(* IEC 61131-3 sources: ArdisCVDCore/codesys/retired_hand_rolled_driver, 11 files *)

(* ---- ST_MfcChannelConfig.st ---- *)
TYPE ST_MfcChannelConfig :
STRUCT
    bSlaveAddr     : BYTE;
    sGasName       : STRING(8);
    rFullScaleSccm : REAL;
END_STRUCT
END_TYPE

(* ---- ST_MfcChannelState.st ---- *)
TYPE ST_MfcChannelState :
STRUCT
    iSubState       : INT;
    iRetryCount     : INT;
    wFaultCode      : WORD;
    xRegulating     : BOOL;
    xFaultActive    : BOOL;
    xCloseConfirmed : BOOL;
    rMeasuredSccm   : REAL;
END_STRUCT
END_TYPE

(* ---- F_MbReadFrame.st ---- *)
FUNCTION F_MbReadFrame : INT
VAR_INPUT
    bAddr : BYTE;
    wReg  : WORD;
END_VAR
VAR_IN_OUT
    aFrame : ARRAY[0..7] OF BYTE;
END_VAR
VAR
    wCrc : WORD;
END_VAR

aFrame[0] := bAddr;
aFrame[1] := BYTE#16#03;
aFrame[2] := WORD_TO_BYTE(SHR(wReg, 8));
aFrame[3] := WORD_TO_BYTE(wReg AND WORD#16#00FF);
aFrame[4] := BYTE#0;
aFrame[5] := BYTE#1;
wCrc := F_ModbusCrc16(iLen := 6, aData := aFrame);
aFrame[6] := WORD_TO_BYTE(wCrc AND WORD#16#00FF);
aFrame[7] := WORD_TO_BYTE(SHR(wCrc, 8));

F_MbReadFrame := 8;

(* ---- F_MbReadStep.st ---- *)
FUNCTION F_MbReadStep : INT
VAR_INPUT
    xReadDone   : BOOL;
    xReadError  : BOOL;
    udiReadSize : UDINT;
END_VAR
VAR_IN_OUT
    xReadExecute    : BOOL;
    xRetriggerArmed : BOOL;
    iRxAccum        : INT;
    iRxIdleScans    : INT;
END_VAR
VAR CONSTANT
    C_MAX_FRAME       : INT := 8;
    C_IDLE_SCAN_LIMIT : INT := 2;
    C_NODATA_LIMIT    : INT := 3;
END_VAR

IF xRetriggerArmed THEN
    xRetriggerArmed := FALSE;
    xReadExecute := TRUE;
    F_MbReadStep := 0;
    RETURN;
END_IF;

IF xReadError THEN
    xReadExecute := FALSE;
    F_MbReadStep := 2;
    RETURN;
END_IF;

IF NOT xReadDone THEN
    F_MbReadStep := 0;
    RETURN;
END_IF;

IF udiReadSize > UDINT#0 THEN
    iRxAccum := iRxAccum + UDINT_TO_INT(udiReadSize);
    iRxIdleScans := 0;
ELSE
    iRxIdleScans := iRxIdleScans + 1;
END_IF;

IF iRxAccum >= C_MAX_FRAME THEN
    xReadExecute := FALSE;
    F_MbReadStep := 1;
    RETURN;
END_IF;

IF (iRxAccum > 0) AND (iRxIdleScans >= C_IDLE_SCAN_LIMIT) THEN
    xReadExecute := FALSE;
    F_MbReadStep := 1;
    RETURN;
END_IF;

IF (iRxAccum = 0) AND (iRxIdleScans >= C_NODATA_LIMIT) THEN
    xReadExecute := FALSE;
    F_MbReadStep := 2;
    RETURN;
END_IF;

xReadExecute := FALSE;
xRetriggerArmed := TRUE;
F_MbReadStep := 0;

(* ---- F_MbRetryOrFault.st ---- *)
FUNCTION F_MbRetryOrFault : INT
VAR_INPUT
    iIssueState : INT;
    iFaultState : INT;
    iMaxRetries : INT;
END_VAR
VAR_IN_OUT
    iRetryCount : INT;
END_VAR

IF iRetryCount < iMaxRetries THEN
    iRetryCount := iRetryCount + 1;
    F_MbRetryOrFault := iIssueState;
ELSE
    iRetryCount := 0;
    F_MbRetryOrFault := iFaultState;
END_IF;

(* ---- F_MbValidateResponse.st ---- *)
FUNCTION F_MbValidateResponse : WORD
VAR_INPUT
    iSize        : INT;
    bExpectAddr  : BYTE;
    bExpectFunc  : BYTE;
    wExpectReg   : WORD;
    wExpectValue : WORD;
    xIsWrite     : BOOL;
END_VAR
VAR_IN_OUT
    aFrame : ARRAY[0..7] OF BYTE;
END_VAR
VAR_OUTPUT
    wReadValue : WORD;
END_VAR
VAR
    wCrcCalc   : WORD;
    wCrcRecv   : WORD;
    iExpectLen : INT;
END_VAR

wReadValue := WORD#0;

IF xIsWrite THEN
    iExpectLen := 8;
ELSE
    iExpectLen := 7;
END_IF;

IF (iSize <> iExpectLen) AND (iSize <> 5) THEN
    F_MbValidateResponse := WORD#5;
    RETURN;
END_IF;

wCrcCalc := F_ModbusCrc16(iLen := iSize - 2, aData := aFrame);
wCrcRecv := BYTE_TO_WORD(aFrame[iSize - 2]) OR SHL(BYTE_TO_WORD(aFrame[iSize - 1]), 8);
IF wCrcCalc <> wCrcRecv THEN
    F_MbValidateResponse := WORD#3;
    RETURN;
END_IF;

IF aFrame[0] <> bExpectAddr THEN
    F_MbValidateResponse := WORD#6;
    RETURN;
END_IF;

IF aFrame[1] = (bExpectFunc OR BYTE#16#80) THEN
    F_MbValidateResponse := WORD#4;
    RETURN;
END_IF;

IF aFrame[1] <> bExpectFunc THEN
    F_MbValidateResponse := WORD#7;
    RETURN;
END_IF;

IF xIsWrite THEN
    IF (aFrame[2] <> WORD_TO_BYTE(SHR(wExpectReg, 8))) OR
       (aFrame[3] <> WORD_TO_BYTE(wExpectReg AND WORD#16#00FF)) OR
       (aFrame[4] <> WORD_TO_BYTE(SHR(wExpectValue, 8))) OR
       (aFrame[5] <> WORD_TO_BYTE(wExpectValue AND WORD#16#00FF)) THEN
        F_MbValidateResponse := WORD#8;
        RETURN;
    END_IF;
ELSE
    wReadValue := SHL(BYTE_TO_WORD(aFrame[3]), 8) OR BYTE_TO_WORD(aFrame[4]);
END_IF;

F_MbValidateResponse := WORD#0;

(* ---- F_MbWriteFrame.st ---- *)
FUNCTION F_MbWriteFrame : INT
VAR_INPUT
    bAddr  : BYTE;
    wReg   : WORD;
    wValue : WORD;
END_VAR
VAR_IN_OUT
    aFrame : ARRAY[0..7] OF BYTE;
END_VAR
VAR
    wCrc : WORD;
END_VAR

aFrame[0] := bAddr;
aFrame[1] := BYTE#16#06;
aFrame[2] := WORD_TO_BYTE(SHR(wReg, 8));
aFrame[3] := WORD_TO_BYTE(wReg AND WORD#16#00FF);
aFrame[4] := WORD_TO_BYTE(SHR(wValue, 8));
aFrame[5] := WORD_TO_BYTE(wValue AND WORD#16#00FF);
wCrc := F_ModbusCrc16(iLen := 6, aData := aFrame);
aFrame[6] := WORD_TO_BYTE(wCrc AND WORD#16#00FF);
aFrame[7] := WORD_TO_BYTE(SHR(wCrc, 8));

F_MbWriteFrame := 8;

(* ---- F_ModbusCrc16.st ---- *)
FUNCTION F_ModbusCrc16 : WORD
VAR_INPUT
    iLen : INT;
END_VAR
VAR_IN_OUT
    aData : ARRAY[0..7] OF BYTE;
END_VAR
VAR
    wCrc : WORD;
    i    : INT;
    j    : INT;
END_VAR

wCrc := WORD#16#FFFF;
FOR i := 0 TO iLen - 1 DO
    wCrc := wCrc XOR BYTE_TO_WORD(aData[i]);
    FOR j := 0 TO 7 DO
        IF (wCrc AND WORD#16#0001) = WORD#16#0001 THEN
            wCrc := SHR(wCrc, 1) XOR WORD#16#A001;
        ELSE
            wCrc := SHR(wCrc, 1);
        END_IF;
    END_FOR;
END_FOR;

F_ModbusCrc16 := wCrc;

(* ---- FB_IncrementalPidOLD.st ---- *)
FUNCTION_BLOCK FB_IncrementalPid
VAR_INPUT
    xEnable       : BOOL;
    xReset        : BOOL;
    xDirectMode   : BOOL;
    rSetpoint     : REAL;
    rMeasured     : REAL;
    rKp           : REAL;
    rKi           : REAL;
    rKd           : REAL;
    rLowerLimit   : REAL;
    rUpperLimit   : REAL;
    rDirectValue  : REAL;
    rFlowCorrection     : REAL := 1.0;
    rPressureCorrection : REAL := 1.0;
    rTotalGasFlow       : REAL := 0.0;
    rCycleSeconds : REAL := 0.2;
END_VAR
VAR_OUTPUT
    rError  : REAL;
    rP      : REAL;
    rI      : REAL;
    rD      : REAL;
    rOutput : REAL;
END_VAR
VAR
    rIntegral      : REAL;
    rPreviousError : REAL;
    xInitialized   : BOOL;
    rMin           : REAL;
    rMax           : REAL;
    rFlowScale     : REAL;
    rPressureScale : REAL;
END_VAR

IF rLowerLimit <= rUpperLimit THEN
    rMin := rLowerLimit;
    rMax := rUpperLimit;
ELSE
    rMin := rUpperLimit;
    rMax := rLowerLimit;
END_IF;

rError := rMeasured - rSetpoint;

IF NOT xEnable THEN
    rP := 0.0;
    rI := 0.0;
    rD := 0.0;
    rOutput := rMin;
    rIntegral := 0.0;
    rPreviousError := rError;
    xInitialized := FALSE;
    RETURN;
END_IF;

IF xReset OR NOT xInitialized THEN
    rIntegral := 0.0;
    rPreviousError := rError;
    rOutput := rMin;
    xInitialized := TRUE;
END_IF;

rP := rKp * rError;

IF rCycleSeconds > 0.001 THEN
    rIntegral := rIntegral + rError * rCycleSeconds;
    rD := rKd * (rError - rPreviousError) / rCycleSeconds;
ELSE
    rD := 0.0;
END_IF;

IF (rFlowCorrection > 0.001) AND (rTotalGasFlow > 50.0) THEN
    IF rTotalGasFlow <= 1100.0 THEN
        rFlowScale := ((rTotalGasFlow - 50.0) / (1100.0 - 50.0)) * (rFlowCorrection - 1.0) + 1.0;
    ELSE
        rFlowScale := rFlowCorrection;
    END_IF;

    IF rFlowScale > 0.001 THEN
        rP := rP / rFlowScale;
        rD := rD / rFlowScale;
    END_IF;
END_IF;

IF (rPressureCorrection > 0.001) AND (rMeasured > 10.0) THEN
    IF rMeasured < 500.0 THEN
        rPressureScale := ((rMeasured - 10.0) / (500.0 - 10.0)) * (rPressureCorrection - 1.0) + 1.0;
    ELSE
        rPressureScale := rPressureCorrection;
    END_IF;

    IF rPressureScale > 0.001 THEN
        rP := rP / rPressureScale;
        rD := rD / rPressureScale;
    END_IF;
END_IF;

IF rIntegral > 1000000.0 THEN
    rIntegral := 1000000.0;
ELSIF rIntegral < -1000000.0 THEN
    rIntegral := -1000000.0;
END_IF;

rI := rKi * rIntegral;
rPreviousError := rError;

IF xDirectMode THEN
    rOutput := rDirectValue;
ELSE
    rOutput := rOutput + rP + rI + rD;
END_IF;

IF rOutput > rMax THEN
    rOutput := rMax;
ELSIF rOutput < rMin THEN
    rOutput := rMin;
END_IF;

(* ---- FB_MfcModbusMaster.st ---- *)
FUNCTION_BLOCK FB_MfcModbusMaster
VAR_INPUT
    xEnable        : BOOL;
    udiPort        : UDINT := 4;
    udiBaudrate    : UDINT := 19200;
    arSetpointSccm : ARRAY[0..5] OF REAL;
END_VAR
VAR_OUTPUT
    xBusOpen         : BOOL;
    udiSweepCounter  : UDINT;
    arMeasuredSccm   : ARRAY[0..5] OF REAL;
    axRegulating     : ARRAY[0..5] OF BOOL;
    axFaultActive    : ARRAY[0..5] OF BOOL;
    axCloseConfirmed : ARRAY[0..5] OF BOOL;
    awFaultCode      : ARRAY[0..5] OF WORD;
END_VAR
VAR CONSTANT
    C_REG_MODE         : WORD := 2;
    C_REG_SETPOINT     : WORD := 4;
    C_REG_MEASURED     : WORD := 5;
    C_REG_RAMPTIME     : WORD := 19;
    C_REG_RAMPSTEP     : WORD := 20;
    C_REG_RAMPEN       : WORD := 21;
    C_MODE_REGULATE    : WORD := 19;
    C_MODE_CLOSE       : WORD := 10;
    C_RAMPTIME_DEFAULT : WORD := 200;
    C_RAMPSTEP_DEFAULT : WORD := 10;
    C_RAMPEN_DEFAULT   : WORD := 1;
    C_FUNC_READ        : BYTE := 16#03;
    C_FUNC_WRITE       : BYTE := 16#06;
    C_MAX_RETRIES      : INT := 2;
    C_OPEN_RETRY_TICKS : UDINT := 40;
    C_IO_TIMEOUT_US    : UDINT := 100000;
END_VAR
VAR
    aCfg        : ARRAY[0..5] OF ST_MfcChannelConfig;
    xConfigInit : BOOL;

    aCh : ARRAY[0..5] OF ST_MfcChannelState;

    iBusState         : INT;
    iChannel          : INT;
    hCom              : CAA.HANDLE;
    udiOpenRetryTicks : UDINT;

    fbOpen  : COM.Open;
    fbWrite : COM.Write;
    fbRead  : COM.Read;
    aParams : ARRAY[1..7] OF COM.PARAMETER;
    xOpenExecute  : BOOL;
    xWriteExecute : BOOL;
    xReadExecute  : BOOL;

    aTx     : ARRAY[0..7] OF BYTE;
    aRx     : ARRAY[0..7] OF BYTE;
    iRxSize : INT;

    iRxAccum         : INT;
    iRxIdleScans     : INT;
    xRxRetriggerArmed: BOOL;
    iRxOffset        : INT;
    iAccumStatus     : INT;

    bPendingAddr    : BYTE;
    wPendingReg     : WORD;
    wPendingValue   : WORD;

    wValidateResult : WORD;
    wReadValue      : WORD;
    rRaw            : REAL;
    iRawSetpoint    : INT;

    i : INT;
END_VAR

IF NOT xConfigInit THEN
    aCfg[0].bSlaveAddr := BYTE#1; aCfg[0].sGasName := 'H2';  aCfg[0].rFullScaleSccm := 1000.0;
    aCfg[1].bSlaveAddr := BYTE#2; aCfg[1].sGasName := 'CH4'; aCfg[1].rFullScaleSccm := 100.0;
    aCfg[2].bSlaveAddr := BYTE#3; aCfg[2].sGasName := 'O2';  aCfg[2].rFullScaleSccm := 50.0;
    aCfg[3].bSlaveAddr := BYTE#4; aCfg[3].sGasName := 'N2';  aCfg[3].rFullScaleSccm := 1000.0;
    aCfg[4].bSlaveAddr := BYTE#5; aCfg[4].sGasName := 'Ar';  aCfg[4].rFullScaleSccm := 10.0;
    aCfg[5].bSlaveAddr := BYTE#6; aCfg[5].sGasName := 'H22'; aCfg[5].rFullScaleSccm := 1000.0;
    xConfigInit := TRUE;
END_IF;

IF NOT xEnable THEN
    FOR i := 0 TO 5 DO
        IF (aCh[i].iSubState <> 900) AND (aCh[i].iSubState <> 901) AND (aCh[i].iSubState <> 902) THEN
            aCh[i].iSubState := 900;
            aCh[i].iRetryCount := 0;
        END_IF;
    END_FOR;
END_IF;

aParams[1].udiParameterId := COM.CAA_Parameter_Constants.udiPort;
aParams[1].udiValue := udiPort;
aParams[2].udiParameterId := COM.CAA_Parameter_Constants.udiBaudrate;
aParams[2].udiValue := udiBaudrate;
aParams[3].udiParameterId := COM.CAA_Parameter_Constants.udiParity;
aParams[3].udiValue := 2;
aParams[4].udiParameterId := COM.CAA_Parameter_Constants.udiStopBits;
aParams[4].udiValue := 0;
aParams[5].udiParameterId := COM.CAA_Parameter_Constants.udiTimeout;
aParams[5].udiValue := 200000;
aParams[6].udiParameterId := COM.CAA_Parameter_Constants.udiByteSize;
aParams[6].udiValue := 8;
aParams[7].udiParameterId := COM.CAA_Parameter_Constants.udiBinary;
aParams[7].udiValue := 1;

CASE iBusState OF

    0:
        xOpenExecute := TRUE;
        xBusOpen := FALSE;
        IF fbOpen.xDone THEN
            hCom := fbOpen.hCom;
            xOpenExecute := FALSE;
            xBusOpen := TRUE;
            iChannel := 0;
            FOR i := 0 TO 5 DO
                IF xEnable THEN
                    aCh[i].iSubState := 100;
                ELSE
                    aCh[i].iSubState := 900;
                END_IF;
                aCh[i].iRetryCount := 0;
            END_FOR;
            iBusState := 10;
        ELSIF fbOpen.xError THEN
            xOpenExecute := FALSE;
            udiOpenRetryTicks := 0;
            iBusState := 5;
        END_IF;

    5:
        xBusOpen := FALSE;
        udiOpenRetryTicks := udiOpenRetryTicks + 1;
        IF udiOpenRetryTicks >= C_OPEN_RETRY_TICKS THEN
            iBusState := 0;
        END_IF;

    10:
        CASE aCh[iChannel].iSubState OF

            100:
                bPendingAddr := aCfg[iChannel].bSlaveAddr;
                wPendingReg := C_REG_RAMPTIME;
                wPendingValue := C_RAMPTIME_DEFAULT;
                F_MbWriteFrame(bAddr := bPendingAddr, wReg := wPendingReg, wValue := wPendingValue, aFrame := aTx);
                xWriteExecute := TRUE;
                aCh[iChannel].iSubState := 101;

            101:
                IF fbWrite.xDone THEN
                    xWriteExecute := FALSE;
                    xReadExecute := TRUE;
                    iRxAccum := 0;
                    iRxIdleScans := 0;
                    xRxRetriggerArmed := FALSE;
                    aCh[iChannel].iSubState := 102;
                ELSIF fbWrite.xError THEN
                    xWriteExecute := FALSE;
                    aCh[iChannel].wFaultCode := WORD#1;
                    aCh[iChannel].iSubState := F_MbRetryOrFault(iIssueState := 100, iFaultState := 900, iMaxRetries := C_MAX_RETRIES, iRetryCount := aCh[iChannel].iRetryCount);
                END_IF;

            102:
                iAccumStatus := F_MbReadStep(xReadDone := fbRead.xDone, xReadError := fbRead.xError, udiReadSize := fbRead.szSize,
                    xReadExecute := xReadExecute, xRetriggerArmed := xRxRetriggerArmed, iRxAccum := iRxAccum, iRxIdleScans := iRxIdleScans);
                IF iAccumStatus = 1 THEN
                    iRxSize := iRxAccum;
                    wValidateResult := F_MbValidateResponse(iSize := iRxSize, bExpectAddr := bPendingAddr, bExpectFunc := C_FUNC_WRITE,
                        wExpectReg := wPendingReg, wExpectValue := wPendingValue, xIsWrite := TRUE, aFrame := aRx, wReadValue => wReadValue);
                    IF wValidateResult = WORD#0 THEN
                        aCh[iChannel].iRetryCount := 0;
                        aCh[iChannel].iSubState := 110;
                    ELSE
                        aCh[iChannel].wFaultCode := wValidateResult;
                        aCh[iChannel].iSubState := F_MbRetryOrFault(iIssueState := 100, iFaultState := 900, iMaxRetries := C_MAX_RETRIES, iRetryCount := aCh[iChannel].iRetryCount);
                    END_IF;
                ELSIF iAccumStatus = 2 THEN
                    aCh[iChannel].wFaultCode := WORD#2;
                    aCh[iChannel].iSubState := F_MbRetryOrFault(iIssueState := 100, iFaultState := 900, iMaxRetries := C_MAX_RETRIES, iRetryCount := aCh[iChannel].iRetryCount);
                END_IF;

            110:
                bPendingAddr := aCfg[iChannel].bSlaveAddr;
                wPendingReg := C_REG_RAMPSTEP;
                wPendingValue := C_RAMPSTEP_DEFAULT;
                F_MbWriteFrame(bAddr := bPendingAddr, wReg := wPendingReg, wValue := wPendingValue, aFrame := aTx);
                xWriteExecute := TRUE;
                aCh[iChannel].iSubState := 111;

            111:
                IF fbWrite.xDone THEN
                    xWriteExecute := FALSE;
                    xReadExecute := TRUE;
                    iRxAccum := 0;
                    iRxIdleScans := 0;
                    xRxRetriggerArmed := FALSE;
                    aCh[iChannel].iSubState := 112;
                ELSIF fbWrite.xError THEN
                    xWriteExecute := FALSE;
                    aCh[iChannel].wFaultCode := WORD#1;
                    aCh[iChannel].iSubState := F_MbRetryOrFault(iIssueState := 110, iFaultState := 900, iMaxRetries := C_MAX_RETRIES, iRetryCount := aCh[iChannel].iRetryCount);
                END_IF;

            112:
                iAccumStatus := F_MbReadStep(xReadDone := fbRead.xDone, xReadError := fbRead.xError, udiReadSize := fbRead.szSize,
                    xReadExecute := xReadExecute, xRetriggerArmed := xRxRetriggerArmed, iRxAccum := iRxAccum, iRxIdleScans := iRxIdleScans);
                IF iAccumStatus = 1 THEN
                    iRxSize := iRxAccum;
                    wValidateResult := F_MbValidateResponse(iSize := iRxSize, bExpectAddr := bPendingAddr, bExpectFunc := C_FUNC_WRITE,
                        wExpectReg := wPendingReg, wExpectValue := wPendingValue, xIsWrite := TRUE, aFrame := aRx, wReadValue => wReadValue);
                    IF wValidateResult = WORD#0 THEN
                        aCh[iChannel].iRetryCount := 0;
                        aCh[iChannel].iSubState := 120;
                    ELSE
                        aCh[iChannel].wFaultCode := wValidateResult;
                        aCh[iChannel].iSubState := F_MbRetryOrFault(iIssueState := 110, iFaultState := 900, iMaxRetries := C_MAX_RETRIES, iRetryCount := aCh[iChannel].iRetryCount);
                    END_IF;
                ELSIF iAccumStatus = 2 THEN
                    aCh[iChannel].wFaultCode := WORD#2;
                    aCh[iChannel].iSubState := F_MbRetryOrFault(iIssueState := 110, iFaultState := 900, iMaxRetries := C_MAX_RETRIES, iRetryCount := aCh[iChannel].iRetryCount);
                END_IF;

            120:
                bPendingAddr := aCfg[iChannel].bSlaveAddr;
                wPendingReg := C_REG_RAMPEN;
                wPendingValue := C_RAMPEN_DEFAULT;
                F_MbWriteFrame(bAddr := bPendingAddr, wReg := wPendingReg, wValue := wPendingValue, aFrame := aTx);
                xWriteExecute := TRUE;
                aCh[iChannel].iSubState := 121;

            121:
                IF fbWrite.xDone THEN
                    xWriteExecute := FALSE;
                    xReadExecute := TRUE;
                    iRxAccum := 0;
                    iRxIdleScans := 0;
                    xRxRetriggerArmed := FALSE;
                    aCh[iChannel].iSubState := 122;
                ELSIF fbWrite.xError THEN
                    xWriteExecute := FALSE;
                    aCh[iChannel].wFaultCode := WORD#1;
                    aCh[iChannel].iSubState := F_MbRetryOrFault(iIssueState := 120, iFaultState := 900, iMaxRetries := C_MAX_RETRIES, iRetryCount := aCh[iChannel].iRetryCount);
                END_IF;

            122:
                iAccumStatus := F_MbReadStep(xReadDone := fbRead.xDone, xReadError := fbRead.xError, udiReadSize := fbRead.szSize,
                    xReadExecute := xReadExecute, xRetriggerArmed := xRxRetriggerArmed, iRxAccum := iRxAccum, iRxIdleScans := iRxIdleScans);
                IF iAccumStatus = 1 THEN
                    iRxSize := iRxAccum;
                    wValidateResult := F_MbValidateResponse(iSize := iRxSize, bExpectAddr := bPendingAddr, bExpectFunc := C_FUNC_WRITE,
                        wExpectReg := wPendingReg, wExpectValue := wPendingValue, xIsWrite := TRUE, aFrame := aRx, wReadValue => wReadValue);
                    IF wValidateResult = WORD#0 THEN
                        aCh[iChannel].iRetryCount := 0;
                        aCh[iChannel].iSubState := 130;
                    ELSE
                        aCh[iChannel].wFaultCode := wValidateResult;
                        aCh[iChannel].iSubState := F_MbRetryOrFault(iIssueState := 120, iFaultState := 900, iMaxRetries := C_MAX_RETRIES, iRetryCount := aCh[iChannel].iRetryCount);
                    END_IF;
                ELSIF iAccumStatus = 2 THEN
                    aCh[iChannel].wFaultCode := WORD#2;
                    aCh[iChannel].iSubState := F_MbRetryOrFault(iIssueState := 120, iFaultState := 900, iMaxRetries := C_MAX_RETRIES, iRetryCount := aCh[iChannel].iRetryCount);
                END_IF;

            130:
                bPendingAddr := aCfg[iChannel].bSlaveAddr;
                wPendingReg := C_REG_MODE;
                wPendingValue := C_MODE_REGULATE;
                F_MbWriteFrame(bAddr := bPendingAddr, wReg := wPendingReg, wValue := wPendingValue, aFrame := aTx);
                xWriteExecute := TRUE;
                aCh[iChannel].iSubState := 131;

            131:
                IF fbWrite.xDone THEN
                    xWriteExecute := FALSE;
                    xReadExecute := TRUE;
                    iRxAccum := 0;
                    iRxIdleScans := 0;
                    xRxRetriggerArmed := FALSE;
                    aCh[iChannel].iSubState := 132;
                ELSIF fbWrite.xError THEN
                    xWriteExecute := FALSE;
                    aCh[iChannel].wFaultCode := WORD#1;
                    aCh[iChannel].iSubState := F_MbRetryOrFault(iIssueState := 130, iFaultState := 900, iMaxRetries := C_MAX_RETRIES, iRetryCount := aCh[iChannel].iRetryCount);
                END_IF;

            132:
                iAccumStatus := F_MbReadStep(xReadDone := fbRead.xDone, xReadError := fbRead.xError, udiReadSize := fbRead.szSize,
                    xReadExecute := xReadExecute, xRetriggerArmed := xRxRetriggerArmed, iRxAccum := iRxAccum, iRxIdleScans := iRxIdleScans);
                IF iAccumStatus = 1 THEN
                    iRxSize := iRxAccum;
                    wValidateResult := F_MbValidateResponse(iSize := iRxSize, bExpectAddr := bPendingAddr, bExpectFunc := C_FUNC_WRITE,
                        wExpectReg := wPendingReg, wExpectValue := wPendingValue, xIsWrite := TRUE, aFrame := aRx, wReadValue => wReadValue);
                    IF wValidateResult = WORD#0 THEN
                        aCh[iChannel].iRetryCount := 0;
                        aCh[iChannel].wFaultCode := WORD#0;
                        aCh[iChannel].xFaultActive := FALSE;
                        aCh[iChannel].xCloseConfirmed := FALSE;
                        aCh[iChannel].xRegulating := TRUE;
                        aCh[iChannel].iSubState := 200;
                    ELSE
                        aCh[iChannel].wFaultCode := wValidateResult;
                        aCh[iChannel].iSubState := F_MbRetryOrFault(iIssueState := 130, iFaultState := 900, iMaxRetries := C_MAX_RETRIES, iRetryCount := aCh[iChannel].iRetryCount);
                    END_IF;
                ELSIF iAccumStatus = 2 THEN
                    aCh[iChannel].wFaultCode := WORD#2;
                    aCh[iChannel].iSubState := F_MbRetryOrFault(iIssueState := 130, iFaultState := 900, iMaxRetries := C_MAX_RETRIES, iRetryCount := aCh[iChannel].iRetryCount);
                END_IF;

            200:
                rRaw := arSetpointSccm[iChannel] / aCfg[iChannel].rFullScaleSccm * 10000.0;
                IF rRaw < 0.0 THEN
                    rRaw := 0.0;
                END_IF;
                iRawSetpoint := REAL_TO_INT(rRaw + 0.5);
                IF iRawSetpoint > 10000 THEN
                    iRawSetpoint := 10000;
                ELSIF iRawSetpoint < 0 THEN
                    iRawSetpoint := 0;
                END_IF;

                bPendingAddr := aCfg[iChannel].bSlaveAddr;
                wPendingReg := C_REG_SETPOINT;
                wPendingValue := INT_TO_WORD(iRawSetpoint);
                F_MbWriteFrame(bAddr := bPendingAddr, wReg := wPendingReg, wValue := wPendingValue, aFrame := aTx);
                xWriteExecute := TRUE;
                aCh[iChannel].iSubState := 201;

            201:
                IF fbWrite.xDone THEN
                    xWriteExecute := FALSE;
                    xReadExecute := TRUE;
                    iRxAccum := 0;
                    iRxIdleScans := 0;
                    xRxRetriggerArmed := FALSE;
                    aCh[iChannel].iSubState := 202;
                ELSIF fbWrite.xError THEN
                    xWriteExecute := FALSE;
                    aCh[iChannel].wFaultCode := WORD#1;
                    aCh[iChannel].iSubState := F_MbRetryOrFault(iIssueState := 200, iFaultState := 900, iMaxRetries := C_MAX_RETRIES, iRetryCount := aCh[iChannel].iRetryCount);
                END_IF;

            202:
                iAccumStatus := F_MbReadStep(xReadDone := fbRead.xDone, xReadError := fbRead.xError, udiReadSize := fbRead.szSize,
                    xReadExecute := xReadExecute, xRetriggerArmed := xRxRetriggerArmed, iRxAccum := iRxAccum, iRxIdleScans := iRxIdleScans);
                IF iAccumStatus = 1 THEN
                    iRxSize := iRxAccum;
                    wValidateResult := F_MbValidateResponse(iSize := iRxSize, bExpectAddr := bPendingAddr, bExpectFunc := C_FUNC_WRITE,
                        wExpectReg := wPendingReg, wExpectValue := wPendingValue, xIsWrite := TRUE, aFrame := aRx, wReadValue => wReadValue);
                    IF wValidateResult = WORD#0 THEN
                        aCh[iChannel].iRetryCount := 0;
                        aCh[iChannel].iSubState := 210;
                    ELSE
                        aCh[iChannel].wFaultCode := wValidateResult;
                        aCh[iChannel].iSubState := F_MbRetryOrFault(iIssueState := 200, iFaultState := 900, iMaxRetries := C_MAX_RETRIES, iRetryCount := aCh[iChannel].iRetryCount);
                    END_IF;
                ELSIF iAccumStatus = 2 THEN
                    aCh[iChannel].wFaultCode := WORD#2;
                    aCh[iChannel].iSubState := F_MbRetryOrFault(iIssueState := 200, iFaultState := 900, iMaxRetries := C_MAX_RETRIES, iRetryCount := aCh[iChannel].iRetryCount);
                END_IF;

            210:
                bPendingAddr := aCfg[iChannel].bSlaveAddr;
                wPendingReg := C_REG_MEASURED;
                F_MbReadFrame(bAddr := bPendingAddr, wReg := wPendingReg, aFrame := aTx);
                xReadExecute := TRUE;
                iRxAccum := 0;
                iRxIdleScans := 0;
                xRxRetriggerArmed := FALSE;
                aCh[iChannel].iSubState := 211;

            211:
                iAccumStatus := F_MbReadStep(xReadDone := fbRead.xDone, xReadError := fbRead.xError, udiReadSize := fbRead.szSize,
                    xReadExecute := xReadExecute, xRetriggerArmed := xRxRetriggerArmed, iRxAccum := iRxAccum, iRxIdleScans := iRxIdleScans);
                IF iAccumStatus = 1 THEN
                    iRxSize := iRxAccum;
                    wValidateResult := F_MbValidateResponse(iSize := iRxSize, bExpectAddr := bPendingAddr, bExpectFunc := C_FUNC_READ,
                        wExpectReg := wPendingReg, wExpectValue := WORD#0, xIsWrite := FALSE, aFrame := aRx, wReadValue => wReadValue);
                    IF wValidateResult = WORD#0 THEN
                        aCh[iChannel].iRetryCount := 0;
                        aCh[iChannel].rMeasuredSccm := UINT_TO_REAL(WORD_TO_UINT(wReadValue)) / 10000.0 * aCfg[iChannel].rFullScaleSccm;
                        aCh[iChannel].iSubState := 200;
                    ELSE
                        aCh[iChannel].wFaultCode := wValidateResult;
                        aCh[iChannel].iSubState := F_MbRetryOrFault(iIssueState := 210, iFaultState := 900, iMaxRetries := C_MAX_RETRIES, iRetryCount := aCh[iChannel].iRetryCount);
                    END_IF;
                    iChannel := (iChannel + 1) MOD 6;
                    IF iChannel = 0 THEN
                        udiSweepCounter := udiSweepCounter + 1;
                    END_IF;
                ELSIF iAccumStatus = 2 THEN
                    aCh[iChannel].wFaultCode := WORD#2;
                    aCh[iChannel].iSubState := F_MbRetryOrFault(iIssueState := 210, iFaultState := 900, iMaxRetries := C_MAX_RETRIES, iRetryCount := aCh[iChannel].iRetryCount);
                    iChannel := (iChannel + 1) MOD 6;
                    IF iChannel = 0 THEN
                        udiSweepCounter := udiSweepCounter + 1;
                    END_IF;
                END_IF;

            900:
                aCh[iChannel].xFaultActive := xEnable;
                aCh[iChannel].xRegulating := FALSE;
                bPendingAddr := aCfg[iChannel].bSlaveAddr;
                wPendingReg := C_REG_MODE;
                wPendingValue := C_MODE_CLOSE;
                F_MbWriteFrame(bAddr := bPendingAddr, wReg := wPendingReg, wValue := wPendingValue, aFrame := aTx);
                xWriteExecute := TRUE;
                aCh[iChannel].iSubState := 901;

            901:
                IF fbWrite.xDone THEN
                    xWriteExecute := FALSE;
                    xReadExecute := TRUE;
                    iRxAccum := 0;
                    iRxIdleScans := 0;
                    xRxRetriggerArmed := FALSE;
                    aCh[iChannel].iSubState := 902;
                ELSIF fbWrite.xError THEN
                    xWriteExecute := FALSE;
                    aCh[iChannel].wFaultCode := WORD#1;
                    aCh[iChannel].iSubState := 900;
                    iChannel := (iChannel + 1) MOD 6;
                    IF iChannel = 0 THEN
                        udiSweepCounter := udiSweepCounter + 1;
                    END_IF;
                END_IF;

            902:
                iAccumStatus := F_MbReadStep(xReadDone := fbRead.xDone, xReadError := fbRead.xError, udiReadSize := fbRead.szSize,
                    xReadExecute := xReadExecute, xRetriggerArmed := xRxRetriggerArmed, iRxAccum := iRxAccum, iRxIdleScans := iRxIdleScans);
                IF iAccumStatus = 1 THEN
                    iRxSize := iRxAccum;
                    wValidateResult := F_MbValidateResponse(iSize := iRxSize, bExpectAddr := bPendingAddr, bExpectFunc := C_FUNC_WRITE,
                        wExpectReg := wPendingReg, wExpectValue := wPendingValue, xIsWrite := TRUE, aFrame := aRx, wReadValue => wReadValue);
                    IF wValidateResult = WORD#0 THEN
                        aCh[iChannel].xCloseConfirmed := TRUE;
                        IF xEnable THEN
                            aCh[iChannel].iSubState := 100;
                            aCh[iChannel].iRetryCount := 0;
                        ELSE
                            aCh[iChannel].iSubState := 900;
                        END_IF;
                    ELSE
                        aCh[iChannel].wFaultCode := wValidateResult;
                        aCh[iChannel].iSubState := 900;
                    END_IF;
                    iChannel := (iChannel + 1) MOD 6;
                    IF iChannel = 0 THEN
                        udiSweepCounter := udiSweepCounter + 1;
                    END_IF;
                ELSIF iAccumStatus = 2 THEN
                    aCh[iChannel].wFaultCode := WORD#2;
                    aCh[iChannel].iSubState := 900;
                    iChannel := (iChannel + 1) MOD 6;
                    IF iChannel = 0 THEN
                        udiSweepCounter := udiSweepCounter + 1;
                    END_IF;
                END_IF;

            ELSE
                aCh[iChannel].iSubState := 900;
        END_CASE;

    ELSE
        iBusState := 0;
END_CASE;

fbOpen(
    xExecute := xOpenExecute,
    usiListLength := 7,
    pParameterList := ADR(aParams));

fbWrite(
    xExecute := xWriteExecute,
    udiTimeOut := C_IO_TIMEOUT_US,
    hCom := hCom,
    pBuffer := ADR(aTx),
    szSize := SIZEOF(aTx));

iRxOffset := iRxAccum;
IF iRxOffset < 0 THEN
    iRxOffset := 0;
ELSIF iRxOffset > 7 THEN
    iRxOffset := 7;
END_IF;

fbRead(
    xExecute := xReadExecute,
    udiTimeOut := C_IO_TIMEOUT_US,
    hCom := hCom,
    pBuffer := ADR(aRx[iRxOffset]),
    szBuffer := SIZEOF(aRx) - INT_TO_UDINT(iRxOffset));

FOR i := 0 TO 5 DO
    arMeasuredSccm[i]   := aCh[i].rMeasuredSccm;
    axRegulating[i]     := aCh[i].xRegulating;
    axFaultActive[i]    := aCh[i].xFaultActive;
    axCloseConfirmed[i] := aCh[i].xCloseConfirmed;
    awFaultCode[i]      := aCh[i].wFaultCode;
END_FOR;

(* ---- PLC_PRG.st ---- *)
    PROGRAM PLC_PRG
    VAR
        xDoBlinkTest : BOOL;
        wBenchMuAo1Output : ARRAY[0..0] OF WORD;

        xTrafficLightGreen  : BOOL;
        xTrafficLightYellow : BOOL;
        xTrafficLightRed    : BOOL;
        wTrafficLightMask   : WORD;

        awMvAi1Value  : ARRAY[0..1] OF WORD;
        awMvAi1Status : ARRAY[0..0] OF WORD;
        uMvAi1Value   : U_DWORD_REAL;
        wMvAi1Status  : WORD;
        xMvAi1Ok      : BOOL;
        rMvAi1Percent : REAL;
        rMvAi1Voltage : REAL;
        rChMeasuredMv : REAL;

        rChamberMuAo1Command : REAL;
        xChamberMuAo1Clamped : BOOL;
        uiChamberMuAo1Command : UINT;

        fbChamber : FB_IncrementalPid;
        fbPlenum  : FB_IncrementalPid;

        xProtocolOk    : BOOL;
        xChamberEnable : BOOL;
        xPlenumEnable  : BOOL;
        xReset         : BOOL;
        udiCycle       : UDINT;

        rChSetpoint : REAL;
        rChMeasured : REAL;
        rChKp       : REAL;
        rChKi       : REAL;
        rChKd       : REAL;
        rChLower    : REAL;
        rChUpper    : REAL;
        rChDirect   : REAL;

        rPlSetpoint : REAL;
        rPlMeasured : REAL;
        rPlKp       : REAL;
        rPlKi       : REAL;
        rPlKd       : REAL;
        rPlLower    : REAL;
        rPlUpper    : REAL;
        rPlDirect   : REAL;
        dwValue     : DWORD;
        xDoBlinkTestEnable : BOOL;
        xBenchMuAo1Enable : BOOL;
        xBenchMuAo1Clamped : BOOL;
        uiBenchMuAo1Command : UINT;
        uiBenchMuAo1Applied : UINT;
        awMvAi1Raw : ARRAY[0..1] OF WORD;
    END_VAR

xProtocolOk := awHolding[0] = WORD#1;
xChamberEnable := xProtocolOk AND (awHolding[1] AND WORD#16#0001) <> WORD#0;
xPlenumEnable := xProtocolOk AND (awHolding[1] AND WORD#16#0002) <> WORD#0;
xReset := (awHolding[1] AND WORD#16#0004) <> WORD#0;
xTrafficLightGreen  := (awHolding[1] AND WORD#16#0010) <> WORD#0;
xTrafficLightYellow := (awHolding[1] AND WORD#16#0020) <> WORD#0;
xTrafficLightRed    := (awHolding[1] AND WORD#16#0040) <> WORD#0;

wTrafficLightMask := WORD#0;
IF xTrafficLightGreen THEN
    wTrafficLightMask := wTrafficLightMask OR WORD#16#0001;
END_IF;
IF xTrafficLightYellow THEN
    wTrafficLightMask := wTrafficLightMask OR WORD#16#0002;
END_IF;
IF xTrafficLightRed THEN
    wTrafficLightMask := wTrafficLightMask OR WORD#16#0004;
END_IF;

rChamberMuAo1Command := fbChamber.rOutput / 10.0;
xChamberMuAo1Clamped := rChamberMuAo1Command > 500.0;

IF xChamberMuAo1Clamped THEN
    uiChamberMuAo1Command := UINT#500;
ELSE
    uiChamberMuAo1Command := REAL_TO_UINT(rChamberMuAo1Command);
END_IF;

wMvAi1Status := awMvAi1Status[0];
xMvAi1Ok := wMvAi1Status = WORD#16#0000;

uMvAi1Value.dwValue := SHL(WORD_TO_DWORD(awMvAi1Value[1]), 16) OR WORD_TO_DWORD(awMvAi1Value[0]);
rMvAi1Percent := uMvAi1Value.rValue;
rMvAi1Voltage := LIMIT(0.0, rMvAi1Percent / 10.0, 10.0);

IF xMvAi1Ok THEN
    rChMeasuredMv := LIMIT(0.0, rMvAi1Percent * 10.0, 1000.0);
END_IF;

rChSetpoint := F_ReadFixed(awHolding[4], awHolding[5]);
rChMeasured := rChMeasuredMv;
rChKp := F_ReadFixed(awHolding[8], awHolding[9]);
rChKi := F_ReadFixed(awHolding[10], awHolding[11]);
rChKd := F_ReadFixed(awHolding[12], awHolding[13]);
rChLower := F_ReadFixed(awHolding[14], awHolding[15]);
rChUpper := F_ReadFixed(awHolding[16], awHolding[17]);
rChDirect := F_ReadFixed(awHolding[18], awHolding[19]);

rPlSetpoint := F_ReadFixed(awHolding[30], awHolding[31]);
rPlMeasured := F_ReadFixed(awHolding[32], awHolding[33]);
rPlKp := F_ReadFixed(awHolding[34], awHolding[35]);
rPlKi := F_ReadFixed(awHolding[36], awHolding[37]);
rPlKd := F_ReadFixed(awHolding[38], awHolding[39]);
rPlLower := F_ReadFixed(awHolding[40], awHolding[41]);
rPlUpper := F_ReadFixed(awHolding[42], awHolding[43]);
rPlDirect := F_ReadFixed(awHolding[44], awHolding[45]);

fbChamber(
    xEnable := xChamberEnable,
    xReset := xReset,
    xDirectMode := awHolding[20] <> WORD#0,
    rSetpoint := rChSetpoint,
    rMeasured := rChMeasured,
    rKp := rChKp,
    rKi := rChKi,
    rKd := rChKd,
    rLowerLimit := rChLower,
    rUpperLimit := rChUpper,
    rDirectValue := rChDirect,
    rCycleSeconds := 0.2);

fbPlenum(
    xEnable := xPlenumEnable,
    xReset := xReset,
    xDirectMode := awHolding[46] <> WORD#0,
    rSetpoint := rPlSetpoint,
    rMeasured := rPlMeasured,
    rKp := rPlKp,
    rKi := rPlKi,
    rKd := rPlKd,
    rLowerLimit := rPlLower,
    rUpperLimit := rPlUpper,
    rDirectValue := rPlDirect,
    rCycleSeconds := 0.2);

udiCycle := udiCycle + 1;
xDoBlinkTestEnable := awHolding[150] = WORD#16#A55A;
xDoBlinkTest := xDoBlinkTestEnable AND ((udiCycle MOD UDINT#10) < UDINT#5);

awHolding[100] := WORD#1;
IF xProtocolOk THEN
    awHolding[101] := WORD#16#0003;
ELSE
    awHolding[101] := WORD#0;
END_IF;
awHolding[102] := DWORD_TO_WORD(udiCycle);
awHolding[103] := DWORD_TO_WORD(SHR(udiCycle, 16));

dwValue := F_ToFixed(fbChamber.rError);
awHolding[104] := DWORD_TO_WORD(dwValue);
awHolding[105] := DWORD_TO_WORD(SHR(dwValue, 16));
dwValue := F_ToFixed(fbChamber.rP);
awHolding[106] := DWORD_TO_WORD(dwValue);
awHolding[107] := DWORD_TO_WORD(SHR(dwValue, 16));
dwValue := F_ToFixed(fbChamber.rI);
awHolding[108] := DWORD_TO_WORD(dwValue);
awHolding[109] := DWORD_TO_WORD(SHR(dwValue, 16));
dwValue := F_ToFixed(fbChamber.rD);
awHolding[110] := DWORD_TO_WORD(dwValue);
awHolding[111] := DWORD_TO_WORD(SHR(dwValue, 16));
dwValue := F_ToFixed(fbChamber.rOutput);
awHolding[112] := DWORD_TO_WORD(dwValue);
awHolding[113] := DWORD_TO_WORD(SHR(dwValue, 16));

dwValue := F_ToFixed(fbPlenum.rError);
awHolding[120] := DWORD_TO_WORD(dwValue);
awHolding[121] := DWORD_TO_WORD(SHR(dwValue, 16));
dwValue := F_ToFixed(fbPlenum.rP);
awHolding[122] := DWORD_TO_WORD(dwValue);
awHolding[123] := DWORD_TO_WORD(SHR(dwValue, 16));
dwValue := F_ToFixed(fbPlenum.rI);
awHolding[124] := DWORD_TO_WORD(dwValue);
awHolding[125] := DWORD_TO_WORD(SHR(dwValue, 16));
dwValue := F_ToFixed(fbPlenum.rD);
awHolding[126] := DWORD_TO_WORD(dwValue);
awHolding[127] := DWORD_TO_WORD(SHR(dwValue, 16));
dwValue := F_ToFixed(fbPlenum.rOutput);
awHolding[128] := DWORD_TO_WORD(dwValue);
awHolding[129] := DWORD_TO_WORD(SHR(dwValue, 16));

dwValue := F_ToFixed(rChMeasuredMv);
awHolding[130] := DWORD_TO_WORD(dwValue);
awHolding[131] := DWORD_TO_WORD(SHR(dwValue, 16));
awHolding[132] := wMvAi1Status;

uiBenchMuAo1Command := WORD_TO_UINT(awHolding[154]);
xBenchMuAo1Enable := awHolding[155] = WORD#16#A55A;
xBenchMuAo1Clamped := uiBenchMuAo1Command > UINT#500;

IF xBenchMuAo1Clamped THEN
    uiBenchMuAo1Command := UINT#500;
END_IF;

IF xBenchMuAo1Enable THEN
    uiBenchMuAo1Applied := uiBenchMuAo1Command;
ELSE
    uiBenchMuAo1Applied := UINT#0;
END_IF;

IF xBenchMuAo1Enable THEN
    awHolding[157] := awHolding[157] OR WORD#16#0001;
END_IF;

IF xBenchMuAo1Clamped THEN
    awHolding[157] := awHolding[157] OR WORD#16#0002;
END_IF;

IF fbChamber.rOutput <= 0.0 THEN
    uiChamberMuAo1Command := UINT#0;
    xChamberMuAo1Clamped := FALSE;
ELSE
    rChamberMuAo1Command := fbChamber.rOutput / 10.0;
    xChamberMuAo1Clamped := rChamberMuAo1Command > 500.0;

    IF xChamberMuAo1Clamped THEN
        uiChamberMuAo1Command := UINT#500;
    ELSE
        uiChamberMuAo1Command := REAL_TO_UINT(rChamberMuAo1Command);
    END_IF;
END_IF;

IF xBenchMuAo1Enable THEN
    uiBenchMuAo1Applied := uiBenchMuAo1Command;
ELSIF xChamberEnable THEN
    uiBenchMuAo1Applied := uiChamberMuAo1Command;
ELSE
    uiBenchMuAo1Applied := UINT#0;
END_IF;

wBenchMuAo1Output[0] := UINT_TO_WORD(uiBenchMuAo1Applied);
awHolding[156] := wBenchMuAo1Output[0];
